(* IEC 61131-3 sources: llm-plc-st-eval/data/processed_definitivo/gpt-4o-2024-08-06/C8/few_shot, 3 files *)

(* ---- ejec_1.st ---- *)
FUNCTION_BLOCK FB_Valvula
VAR_INPUT
    nivelAlto : BOOL; (* Contacto NA para activar el temporizador *)
END_VAR
VAR_OUTPUT
    valvula : BOOL; (* Bobina controlada por el temporizador *)
END_VAR
VAR
    T1 : TON; (* Temporizador TON *)
END_VAR

(* Configuración del temporizador *)
T1(IN := nivelAlto, PT := T#5S);

(* La salida del temporizador controla la bobina *)
valvula := T1.Q;
END_FUNCTION_BLOCK

(* ---- ejec_2.st ---- *)
FUNCTION_BLOCK FB_Valvula
VAR_INPUT
    nivelAlto : BOOL; (* Contacto NA para activar el temporizador *)
END_VAR
VAR_OUTPUT
    valvula : BOOL; (* Bobina controlada por la salida del temporizador *)
END_VAR
VAR
    T1 : TON; (* Temporizador TON *)
END_VAR

(* Configuración del temporizador TON *)
T1(IN := nivelAlto, PT := T#5S);

(* La salida de la válvula se activa cuando el temporizador alcanza el tiempo preestablecido *)
valvula := T1.Q;
END_FUNCTION_BLOCK

(* ---- ejec_3.st ---- *)
FUNCTION_BLOCK FB_Valvula
VAR_INPUT
    nivelAlto : BOOL; (* Contacto NA que activa el temporizador *)
END_VAR
VAR_OUTPUT
    valvula : BOOL; (* Bobina activada por la salida del temporizador *)
END_VAR
VAR
    T1 : TON; (* Temporizador TON *)
END_VAR

(* Configuración del temporizador TON *)
T1(IN := nivelAlto, PT := T#5S);

(* La salida del temporizador activa la bobina *)
valvula := T1.Q;
END_FUNCTION_BLOCK
